(* IEC 61131-3 sources: SafePLC-Gen-Evaluation/Evaluation Results/Dexpi_PDF/run_05, 2 files *)

(* ---- io_declarations.st ---- *)
(* ==================================================  *)
(* PLC I/O Variable Declarations — CODESYS 3.5  *)
(* Generated by SafePLC-Gen Multimodal  *)
(* ==================================================  *)

VAR_GLOBAL
    (* --- Analog Inputs ---  *)
    PI_4712.01_Raw               AT %IW0       : INT := 0;    (* PI-4712.01 — Pressure indicator PI 4712.01. Local pre  *)
    (* --- Analog Outputs ---  *)
    FC_VALVE_H_1007_Out          AT %QW0       : INT := 0;    (* FC-VALVE-H-1007 — Fail-closed (F.C.) control valve on inle  *)
    PVA_4712.02_Out              AT %QW2       : INT := 0;    (* PVA-4712.02 — Pressure control valve on recirculation   *)
    TV_4750.03_Out               AT %QW4       : INT := 0;    (* TV-4750.03 — Temperature control valve on utility lin  *)
    (* --- Digital Inputs ---  *)
    HS_4750.01                   AT %IX0.0     : BOOL := FALSE;    (* HS-4750.01 — Hand switch HS 4750.01. Located near pum  *)
END_VAR

(* ---- generated_code.st ---- *)
(* Generated by SafePLC-Gen Multimodal — CODESYS 3.5 *)
(* IEC 61131-3 Structured Text *)
(* Date: 2026-04-25T14:06:03.708277 *)

PROGRAM SafePLC_Main

VAR
    PI_4712_01_Raw               AT %IW0       : INT := 0;
    FC_VALVE_H_1007_Out          AT %QW0       : INT := 0;
    PVA_4712_02_Out              AT %QW2       : INT := 0;
    TV_4750_03_Out               AT %QW4       : INT := 0;
    HS_4750_01                   AT %IX0.0     : BOOL := FALSE;
    ESTOP                        AT %IX0.1     : BOOL := FALSE;
    MANUAL_RESET                 AT %IX0.2     : BOOL := FALSE;
END_VAR

VAR
    PI_4712_01_Scaled            : REAL := 0.0;

    PI_4712_01_HH_SP             : REAL := 180.0;
    PI_4712_01_H_SP              : REAL := 160.0;
    PI_4712_01_L_SP              : REAL := 20.0;
    PI_4712_01_LL_SP             : REAL := 10.0;
    PI_4712_01_Deadband          : REAL := 2.0;
    PI_4712_01_H                 : BOOL := FALSE;
    PI_4712_01_L                 : BOOL := FALSE;
    PI_4712_01_HH_Latch          : SR := (S1 := FALSE, R := FALSE, Q1 := FALSE);
    PI_4712_01_LL_Latch          : SR := (S1 := FALSE, R := FALSE, Q1 := FALSE);
    PI_4712_01_HH_Ack            : BOOL := FALSE;
    PI_4712_01_LL_Ack            : BOOL := FALSE;

    LOOP_4750_03_TRIP            : BOOL := FALSE;
    LOOP_4712_02_TRIP            : BOOL := FALSE;
    LOOP_104_01_TRIP             : BOOL := FALSE;

    TICSA_4750_03_HH             : BOOL := FALSE;
    TICSA_4750_03_LL             : BOOL := FALSE;
    PICSA_4712_02_HH             : BOOL := FALSE;
    PICSA_4712_02_LL             : BOOL := FALSE;
    SV_104_01_HH                 : BOOL := FALSE;
    SV_104_01_LL                 : BOOL := FALSE;

    SAFE_STATE                   : BOOL := FALSE;

    TV_4750_03_SP                : REAL := 80.0;
    TV_4750_03_Kp                : REAL := 1.2;
    TV_4750_03_Ki                : REAL := 0.05;
    TV_4750_03_Integral          : REAL := 0.0;
    TV_4750_03_Error             : REAL := 0.0;
    TV_4750_03_Output_Pct        : REAL := 0.0;

    PVA_4712_02_SP               : REAL := 100.0;
    PVA_4712_02_Kp               : REAL := 1.0;
    PVA_4712_02_Ki               : REAL := 0.04;
    PVA_4712_02_Integral         : REAL := 0.0;
    PVA_4712_02_Error            : REAL := 0.0;
    PVA_4712_02_Output_Pct       : REAL := 0.0;

    FC_1007_SP                   : REAL := 50.0;
    FC_1007_Kp                   : REAL := 0.8;
    FC_1007_Ki                   : REAL := 0.03;
    FC_1007_Integral             : REAL := 0.0;
    FC_1007_Error                : REAL := 0.0;
    FC_1007_Output_Pct           : REAL := 0.0;

    SV_104_01_Out                : BOOL := FALSE;
    CHECK_75SA21_Out             : BOOL := FALSE;
    CHECK_P_4711_Out             : BOOL := FALSE;
    BV_73KH12_50_1_Out           : BOOL := FALSE;
    BV_73KH12_50_2_Out           : BOOL := FALSE;
    BV_73KH12_25_1_Out           : BOOL := FALSE;
    BV_73KH12_25_2_Out           : BOOL := FALSE;
    BV_MNc_47125_N5_Out          : BOOL := FALSE;
    BV_MNc_47125_73HG12_Out      : BOOL := FALSE;
    BV_MNc_47127_Q80_Out         : BOOL := FALSE;

    System_Alarm                 : BOOL := FALSE;
    FirstScan                    : BOOL := TRUE;
END_VAR

IF FirstScan THEN
    LOOP_4750_03_TRIP   := TRUE;
    LOOP_4712_02_TRIP   := TRUE;
    LOOP_104_01_TRIP    := TRUE;
    SAFE_STATE          := TRUE;
    TV_4750_03_Out      := 6554;
    PVA_4712_02_Out     := 6554;
    FC_VALVE_H_1007_Out := 6554;
    SV_104_01_Out       := FALSE;
    FirstScan           := FALSE;
    RETURN;
END_IF;

PI_4712_01_Scaled := ((INT_TO_REAL(PI_4712_01_Raw) - 6554.0) /
                      (32767.0 - 6554.0)) * 200.0;

IF PI_4712_01_Scaled >= PI_4712_01_HH_SP THEN
    PI_4712_01_HH_Latch.S1 := TRUE;
ELSIF PI_4712_01_Scaled <= (PI_4712_01_HH_SP - PI_4712_01_Deadband) THEN
    PI_4712_01_HH_Latch.S1 := FALSE;
END_IF;
PI_4712_01_HH_Latch.R := PI_4712_01_HH_Ack AND NOT (PI_4712_01_Scaled >= PI_4712_01_HH_SP);
PI_4712_01_HH_Latch(S1 := PI_4712_01_HH_Latch.S1, R := PI_4712_01_HH_Latch.R);

IF PI_4712_01_Scaled >= PI_4712_01_H_SP THEN
    PI_4712_01_H := TRUE;
ELSIF PI_4712_01_Scaled <= (PI_4712_01_H_SP - PI_4712_01_Deadband) THEN
    PI_4712_01_H := FALSE;
END_IF;

IF PI_4712_01_Scaled <= PI_4712_01_L_SP THEN
    PI_4712_01_L := TRUE;
ELSIF PI_4712_01_Scaled >= (PI_4712_01_L_SP + PI_4712_01_Deadband) THEN
    PI_4712_01_L := FALSE;
END_IF;

IF PI_4712_01_Scaled <= PI_4712_01_LL_SP THEN
    PI_4712_01_LL_Latch.S1 := TRUE;
ELSIF PI_4712_01_Scaled >= (PI_4712_01_LL_SP + PI_4712_01_Deadband) THEN
    PI_4712_01_LL_Latch.S1 := FALSE;
END_IF;
PI_4712_01_LL_Latch.R := PI_4712_01_LL_Ack AND NOT (PI_4712_01_Scaled <= PI_4712_01_LL_SP);
PI_4712_01_LL_Latch(S1 := PI_4712_01_LL_Latch.S1, R := PI_4712_01_LL_Latch.R);

PICSA_4712_02_HH := PI_4712_01_HH_Latch.Q1;
PICSA_4712_02_LL := PI_4712_01_LL_Latch.Q1;

TICSA_4750_03_HH := HS_4750_01;
TICSA_4750_03_LL := FALSE;
SV_104_01_HH     := FALSE;
SV_104_01_LL     := FALSE;

IF TICSA_4750_03_HH OR TICSA_4750_03_LL THEN
    LOOP_4750_03_TRIP := TRUE;
ELSIF LOOP_4750_03_TRIP AND MANUAL_RESET
      AND NOT TICSA_4750_03_HH AND NOT TICSA_4750_03_LL THEN
    LOOP_4750_03_TRIP := FALSE;
END_IF;

IF PICSA_4712_02_HH OR PICSA_4712_02_LL THEN
    LOOP_4712_02_TRIP := TRUE;
ELSIF LOOP_4712_02_TRIP AND MANUAL_RESET
      AND NOT PICSA_4712_02_HH AND NOT PICSA_4712_02_LL THEN
    LOOP_4712_02_TRIP := FALSE;
END_IF;

IF SV_104_01_HH OR SV_104_01_LL THEN
    LOOP_104_01_TRIP := TRUE;
ELSIF LOOP_104_01_TRIP AND MANUAL_RESET
      AND NOT SV_104_01_HH AND NOT SV_104_01_LL THEN
    LOOP_104_01_TRIP := FALSE;
END_IF;

SAFE_STATE := ESTOP
              OR LOOP_4750_03_TRIP
              OR LOOP_4712_02_TRIP
              OR LOOP_104_01_TRIP;

IF NOT SAFE_STATE THEN

    TV_4750_03_Error    := TV_4750_03_SP - PI_4712_01_Scaled;
    TV_4750_03_Integral := TV_4750_03_Integral + (TV_4750_03_Ki * TV_4750_03_Error);
    IF TV_4750_03_Integral > 100.0 THEN
        TV_4750_03_Integral := 100.0;
    ELSIF TV_4750_03_Integral < 0.0 THEN
        TV_4750_03_Integral := 0.0;
    END_IF;
    TV_4750_03_Output_Pct := (TV_4750_03_Kp * TV_4750_03_Error) + TV_4750_03_Integral;
    IF TV_4750_03_Output_Pct > 100.0 THEN
        TV_4750_03_Output_Pct := 100.0;
    ELSIF TV_4750_03_Output_Pct < 0.0 THEN
        TV_4750_03_Output_Pct := 0.0;
    END_IF;
    TV_4750_03_Out := REAL_TO_INT(6554.0 + (TV_4750_03_Output_Pct / 100.0) * (32767.0 - 6554.0));

    PVA_4712_02_Error    := PVA_4712_02_SP - PI_4712_01_Scaled;
    PVA_4712_02_Integral := PVA_4712_02_Integral + (PVA_4712_02_Ki * PVA_4712_02_Error);
    IF PVA_4712_02_Integral > 100.0 THEN
        PVA_4712_02_Integral := 100.0;
    ELSIF PVA_4712_02_Integral < 0.0 THEN
        PVA_4712_02_Integral := 0.0;
    END_IF;
    PVA_4712_02_Output_Pct := (PVA_4712_02_Kp * PVA_4712_02_Error) + PVA_4712_02_Integral;
    IF PVA_4712_02_Output_Pct > 100.0 THEN
        PVA_4712_02_Output_Pct := 100.0;
    ELSIF PVA_4712_02_Output_Pct < 0.0 THEN
        PVA_4712_02_Output_Pct := 0.0;
    END_IF;
    PVA_4712_02_Out := REAL_TO_INT(6554.0 + (PVA_4712_02_Output_Pct / 100.0) * (32767.0 - 6554.0));

    FC_1007_Error    := FC_1007_SP - PI_4712_01_Scaled;
    FC_1007_Integral := FC_1007_Integral + (FC_1007_Ki * FC_1007_Error);
    IF FC_1007_Integral > 100.0 THEN
        FC_1007_Integral := 100.0;
    ELSIF FC_1007_Integral < 0.0 THEN
        FC_1007_Integral := 0.0;
    END_IF;
    FC_1007_Output_Pct := (FC_1007_Kp * FC_1007_Error) + FC_1007_Integral;
    IF FC_1007_Output_Pct > 100.0 THEN
        FC_1007_Output_Pct := 100.0;
    ELSIF FC_1007_Output_Pct < 0.0 THEN
        FC_1007_Output_Pct := 0.0;
    END_IF;
    FC_VALVE_H_1007_Out := REAL_TO_INT(6554.0 + (FC_1007_Output_Pct / 100.0) * (32767.0 - 6554.0));

    SV_104_01_Out           := NOT HS_4750_01;
    CHECK_75SA21_Out        := TRUE;
    CHECK_P_4711_Out        := TRUE;
    BV_73KH12_50_1_Out      := TRUE;
    BV_73KH12_50_2_Out      := TRUE;
    BV_73KH12_25_1_Out      := TRUE;
    BV_73KH12_25_2_Out      := TRUE;
    BV_MNc_47125_N5_Out     := TRUE;
    BV_MNc_47125_73HG12_Out := TRUE;
    BV_MNc_47127_Q80_Out    := TRUE;

ELSE
    TV_4750_03_Out          := 6554;
    PVA_4712_02_Out         := 6554;
    FC_VALVE_H_1007_Out     := 6554;
    SV_104_01_Out           := FALSE;
    CHECK_75SA21_Out        := FALSE;
    CHECK_P_4711_Out        := FALSE;
    BV_73KH12_50_1_Out      := FALSE;
    BV_73KH12_50_2_Out      := FALSE;
    BV_73KH12_25_1_Out      := FALSE;
    BV_73KH12_25_2_Out      := FALSE;
    BV_MNc_47125_N5_Out     := FALSE;
    BV_MNc_47125_73HG12_Out := FALSE;
    BV_MNc_47127_Q80_Out    := FALSE;
    TV_4750_03_Integral     := 0.0;
    PVA_4712_02_Integral    := 0.0;
    FC_1007_Integral        := 0.0;
END_IF;

System_Alarm :=
    PI_4712_01_HH_Latch.Q1 OR PI_4712_01_LL_Latch.Q1 OR
    PI_4712_01_H            OR PI_4712_01_L            OR
    LOOP_4750_03_TRIP       OR LOOP_4712_02_TRIP        OR
    LOOP_104_01_TRIP        OR SAFE_STATE;

END_PROGRAM
